// TIA Portal project "Clase2_PLCN3y4" (V13)

(* hardware
DEVICE "S7-1200 station_1"  S7-1200 Station
   slot 0: "Rack_0"  Rack  V1.0
   slot 1: "PLC_1"  CPU 1214C AC/DC/Rly  6ES7 214-1BE30-0XB0  V2.2
*)

// ===== PLC "PLC_1"  CPU 1214C AC/DC/Rly =====

VAR_GLOBAL   // PLC tag table "Tabla de variables estándar"
   "inicio" AT %I0.0 : Bool;
   "mem1" AT %M10.0 : Bool;
   "salida" AT %Q0.0 : Bool;
   "value" AT %IW64 : UInt;
   "norm" AT %MD100 : Real;
   "scale" AT %MD120 : DWord;
   "t_conv" AT %MD200 : DWord;
   "t_out" AT %MD220 : DWord;
END_VAR

// folder: System blocks/Program resources

DATA_BLOCK "TEM1"   // DB1
{ S7_Optimized_Access := 'FALSE' }
AUTHOR : Simatic
FAMILY : IEC
NAME : IEC_TMR
VERSION : 1.0
// stored: InstanceOfName ?
"?"
BEGIN
END_DATA_BLOCK

// folder: (top level)

ORGANIZATION_BLOCK "Main"   // OB1, LAD, ProgramCycle
TITLE = "Main Program Sweep (Cycle)"
{ S7_Optimized_Access := 'FALSE' }
VERSION : 0.1
// S
BEGIN

REGION Network 1
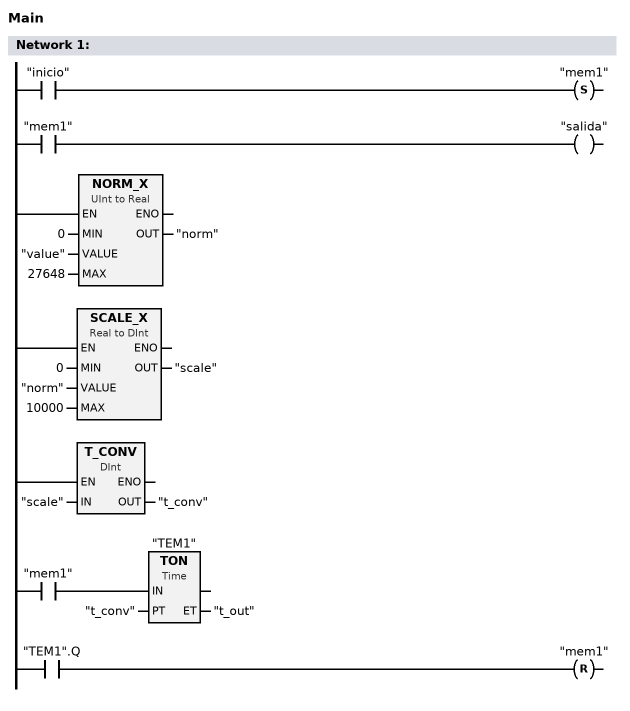
   IF "inicio" THEN "mem1" := TRUE; END_IF;
   "salida" := "mem1";
   "norm" := NORM_X(MIN := 0, VALUE := "value", MAX := 27648);
   "scale" := SCALE_X(MIN := 0, VALUE := "norm", MAX := 10000);
   "t_conv" := T_CONV(IN := "scale");
   "TEM1".TON(IN := "mem1", PT := "t_conv", ET => "t_out");
   IF "TEM1".Q THEN "mem1" := FALSE; END_IF;
END_REGION
END_ORGANIZATION_BLOCK